(* Logix 5000 project; controller R400_500_XLS vendor 1 type 14 code 216 rev 31.11; software revision 31.01; part 22 of 32 *)
(* tags used below, declared in another part *)
   Abort1 : DINT;   // Not Used
   Alarm : SINT;   // Wait 3 seconds
   AlarmAcked : BOOL;   // Alarm has been acked
   bAlrm : BOOL[64];
   CycExcBuffer : UDT_CYCLE;
   CycleSequence : UDT_CYCLE_SEQUENCE;
   DrnSmp : DINT;
   DRYING : DINT;   // Drying id number
   F1rinse : DINT;   // Not Used
   F2rinse : DINT;   // Not Used
   F3rinse : DINT;   // Not Used
   F4rinse : INT;   // Transition for the conductivity based evalutaion
   F4rinse_Tran : INT;   // Transitions for the conductivity based evaluation
   FINAL_RINSE_MAX_NBR : INT;   // Maximum nimber of final rinse
   M : DINT[5];   // Memory Bits
   NbFinalRinseDone : DINT;
   ONS_FC08 : DINT;
   Run : DINT;
   SumpWaterVolume : DINT;   // Sump Water Volume 0 =Low 1= High
   Tmr : TIMER[107];
   WaterSaved : BOOL;   // Water Saved In Sump (Last Final Rinse Water)
   ENABLE : BOOL;   // Enable bit
   FinalRinseCond : REAL;
   I_Pw_Tnk_Lvl_Sw : BOOL;   // Pure water tank level switch
   TreatmentPtr : DINT;
   Unit : Hrdwre;   // Unit Configuration
(* MainProgram, continued *)

ROUTINE WSH_16_TRT_FRINSE   (* ladder *)
// This routine performs the Final Rinse treatments
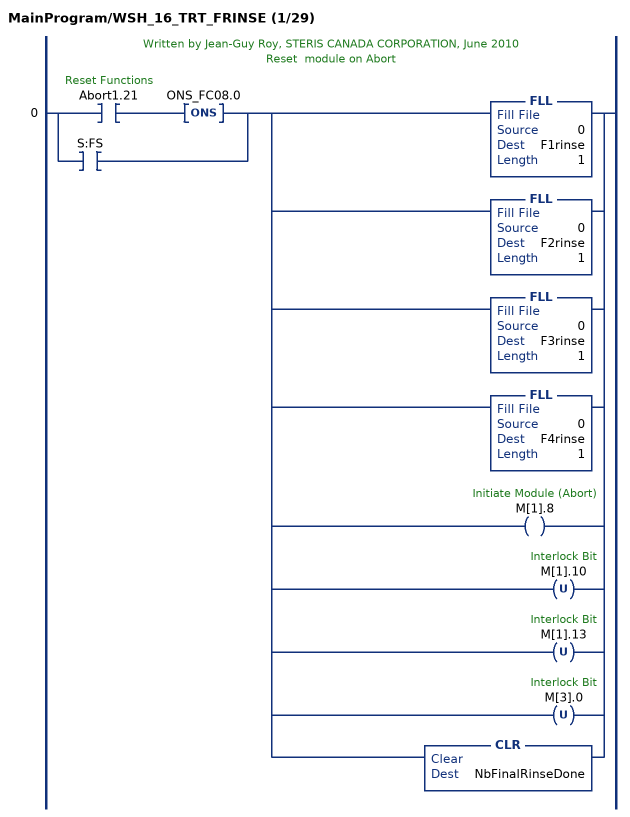
   // Written by Jean-Guy Roy, STERIS CANADA CORPORATION, June 2010
   // Reset  module on Abort
   0: [XIC(Abort1.21) ONS(ONS_FC08.0) ,XIC(S:FS) ][FLL(0,F1rinse,1) ,FLL(0,F2rinse,1) ,FLL(0,F3rinse,1) ,FLL(0,F4rinse,1) ,OTE(M[1].8) ,OTU(M[1].10) ,OTU(M[1].13) ,OTU(M[3].0) ,CLR(NbFinalRinseDone) ];
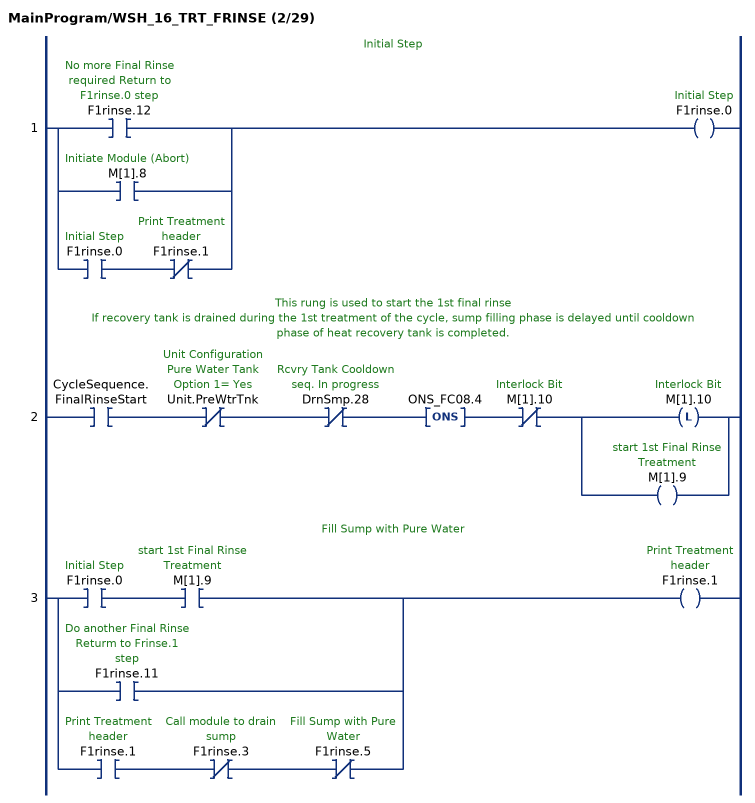
   // Initial Step
   1: [XIC(F1rinse.12) ,XIC(M[1].8) ,XIC(F1rinse.0) XIO(F1rinse.1) ]OTE(F1rinse.0);
   // This rung is used to start the 1st final rinse
   // If recovery tank is drained during the 1st treatment of the cycle, sump filling phase is delayed until cooldown phase of heat recovery tank is completed.
   2: XIC(CycleSequence.FinalRinseStart)XIO(Unit.PreWtrTnk)XIO(DrnSmp.28)ONS(ONS_FC08.4)XIO(M[1].10)[OTL(M[1].10) ,OTE(M[1].9) ];
   // Fill Sump with Pure Water
   3: [XIC(F1rinse.0) XIC(M[1].9) ,XIC(F1rinse.11) ,XIC(F1rinse.1) XIO(F1rinse.3) XIO(F1rinse.5) ]OTE(F1rinse.1);
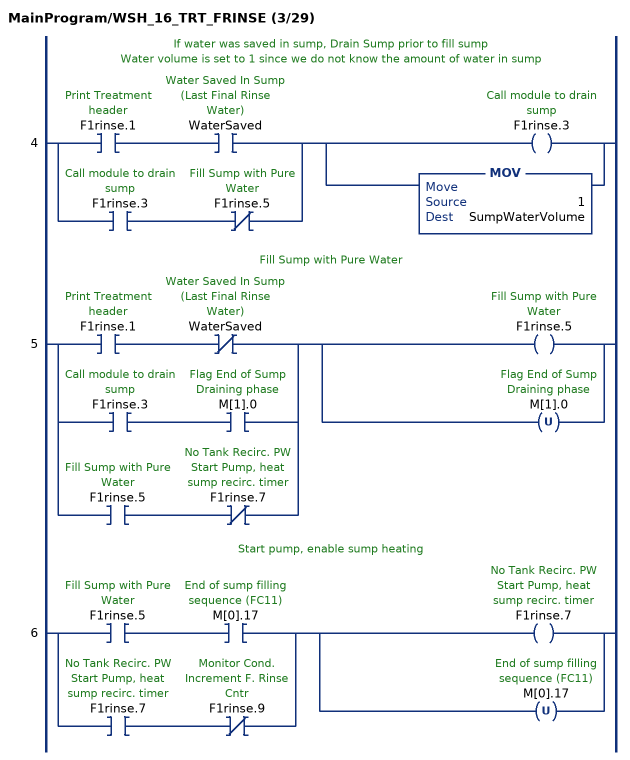
   // If water was saved in sump, Drain Sump prior to fill sump
   // Water volume is set to 1 since we do not know the amount of water in sump
   4: [XIC(F1rinse.1) XIC(WaterSaved) ,XIC(F1rinse.3) XIO(F1rinse.5) ][OTE(F1rinse.3) ,MOV(1,SumpWaterVolume) ];
   // Fill Sump with Pure Water
   5: [[XIC(F1rinse.1) XIO(WaterSaved) ,XIC(F1rinse.3) XIC(M[1].0) ] ,XIC(F1rinse.5) XIO(F1rinse.7) ][OTE(F1rinse.5) ,OTU(M[1].0) ];
   // Start pump, enable sump heating
   6: [XIC(F1rinse.5) XIC(M[0].17) ,XIC(F1rinse.7) XIO(F1rinse.9) ][OTE(F1rinse.7) ,OTU(M[0].17) ];
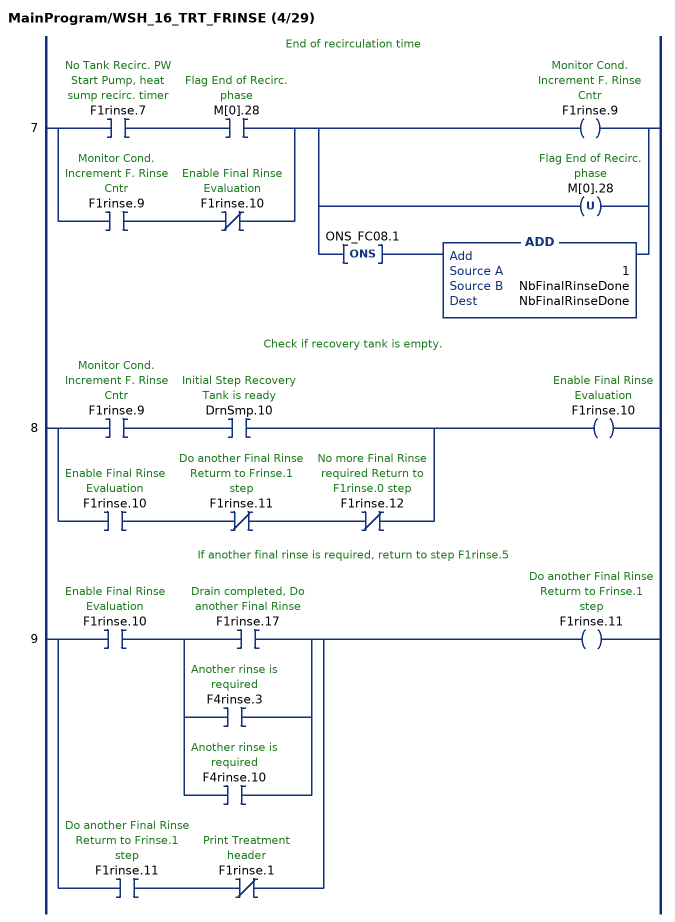
   // End of recirculation time
   7: [XIC(F1rinse.7) XIC(M[0].28) ,XIC(F1rinse.9) XIO(F1rinse.10) ][[OTE(F1rinse.9) ,OTU(M[0].28) ] ,ONS(ONS_FC08.1) ADD(1,NbFinalRinseDone,NbFinalRinseDone) ];
   // Check if recovery tank is empty.
   8: [XIC(F1rinse.9) XIC(DrnSmp.10) ,XIC(F1rinse.10) XIO(F1rinse.11) XIO(F1rinse.12) ]OTE(F1rinse.10);
   // If another final rinse is required, return to step F1rinse.5
   9: [XIC(F1rinse.10) [XIC(F1rinse.17) ,XIC(F4rinse.3) ,XIC(F4rinse.10) ] ,XIC(F1rinse.11) XIO(F1rinse.1) ]OTE(F1rinse.11);
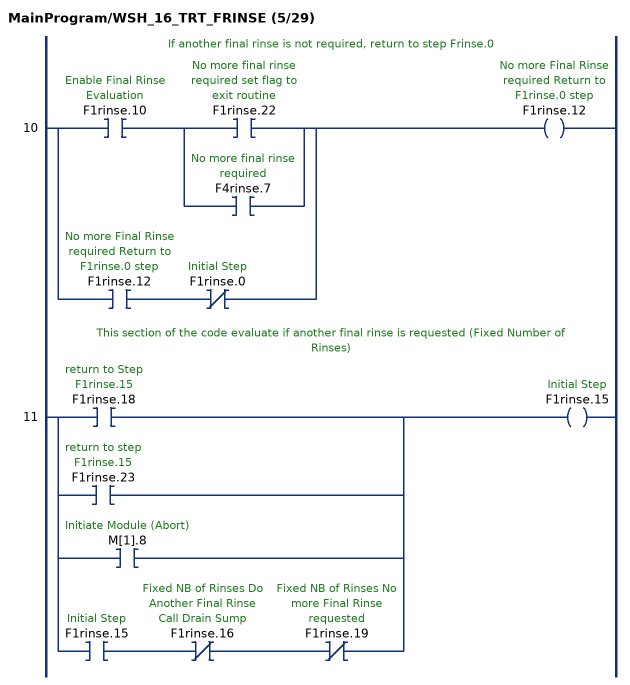
   // If another final rinse is not required, return to step Frinse.0
   10: [XIC(F1rinse.10) [XIC(F1rinse.22) ,XIC(F4rinse.7) ] ,XIC(F1rinse.12) XIO(F1rinse.0) ]OTE(F1rinse.12);
   // This section of the code evaluate if another final rinse is requested (Fixed Number of Rinses)
   11: [XIC(F1rinse.18) ,XIC(F1rinse.23) ,XIC(M[1].8) ,XIC(F1rinse.15) XIO(F1rinse.16) XIO(F1rinse.19) ]OTE(F1rinse.15);
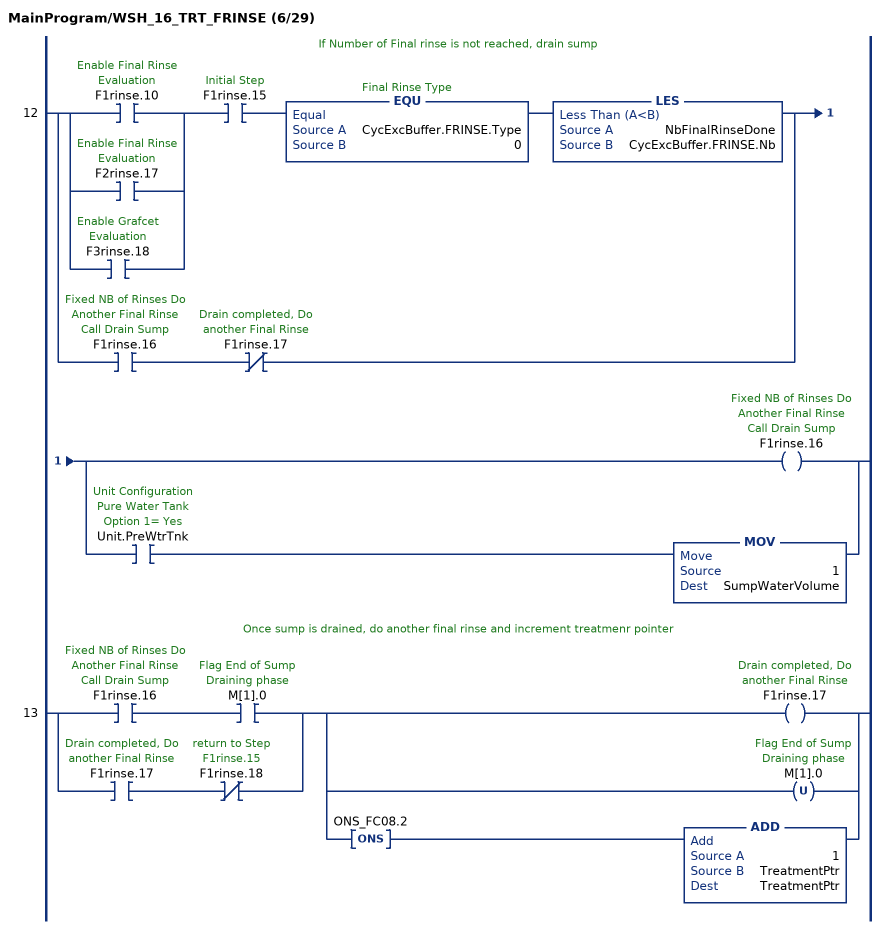
   // If Number of Final rinse is not reached, drain sump
   12: [[XIC(F1rinse.10) ,XIC(F2rinse.17) ,XIC(F3rinse.18) ] XIC(F1rinse.15) EQU(CycExcBuffer.FRINSE.Type,0) LES(NbFinalRinseDone,CycExcBuffer.FRINSE.Nb) ,XIC(F1rinse.16) XIO(F1rinse.17) ][OTE(F1rinse.16) ,XIC(Unit.PreWtrTnk) MOV(1,SumpWaterVolume) ];
   // Once sump is drained, do another final rinse and increment treatmenr pointer
   13: [XIC(F1rinse.16) XIC(M[1].0) ,XIC(F1rinse.17) XIO(F1rinse.18) ][OTE(F1rinse.17) ,OTU(M[1].0) ,ONS(ONS_FC08.2) ADD(1,TreatmentPtr,TreatmentPtr) ];
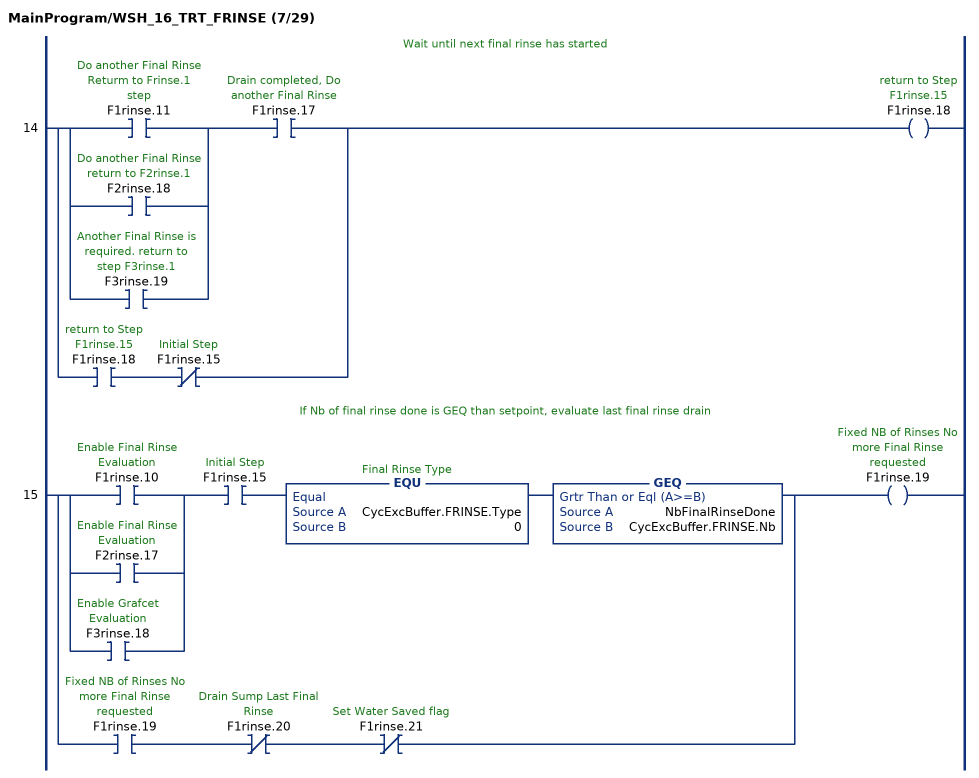
   // Wait until next final rinse has started
   14: [[XIC(F1rinse.11) ,XIC(F2rinse.18) ,XIC(F3rinse.19) ] XIC(F1rinse.17) ,XIC(F1rinse.18) XIO(F1rinse.15) ]OTE(F1rinse.18);
   // If Nb of final rinse done is GEQ than setpoint, evaluate last final rinse drain
   15: [[XIC(F1rinse.10) ,XIC(F2rinse.17) ,XIC(F3rinse.18) ] XIC(F1rinse.15) EQU(CycExcBuffer.FRINSE.Type,0) GEQ(NbFinalRinseDone,CycExcBuffer.FRINSE.Nb) ,XIC(F1rinse.19) XIO(F1rinse.20) XIO(F1rinse.21) ]OTE(F1rinse.19);
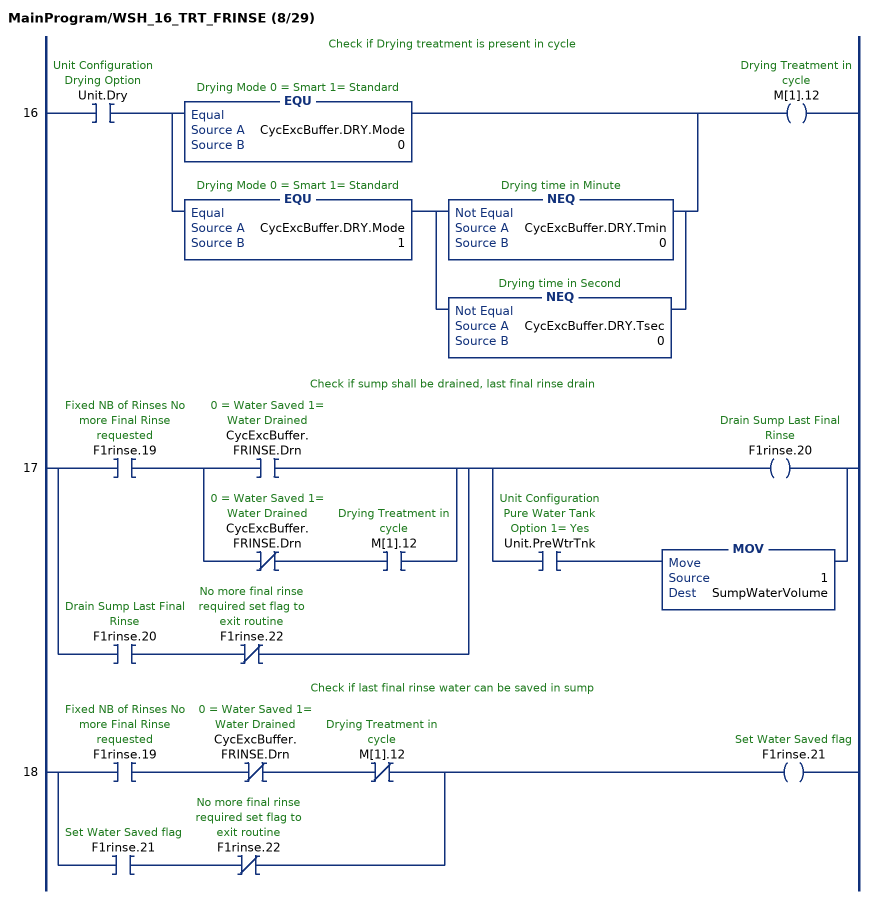
   // Check if Drying treatment is present in cycle
   16: XIC(Unit.Dry)[EQU(CycExcBuffer.DRY.Mode,0) ,EQU(CycExcBuffer.DRY.Mode,1) [NEQ(CycExcBuffer.DRY.Tmin,0) ,NEQ(CycExcBuffer.DRY.Tsec,0) ] ]OTE(M[1].12);
   // Check if sump shall be drained, last final rinse drain
   17: [XIC(F1rinse.19) [XIC(CycExcBuffer.FRINSE.Drn) ,XIO(CycExcBuffer.FRINSE.Drn) XIC(M[1].12) ] ,XIC(F1rinse.20) XIO(F1rinse.22) ][OTE(F1rinse.20) ,XIC(Unit.PreWtrTnk) MOV(1,SumpWaterVolume) ];
   // Check if last final rinse water can be saved in sump
   18: [XIC(F1rinse.19) XIO(CycExcBuffer.FRINSE.Drn) XIO(M[1].12) ,XIC(F1rinse.21) XIO(F1rinse.22) ]OTE(F1rinse.21);
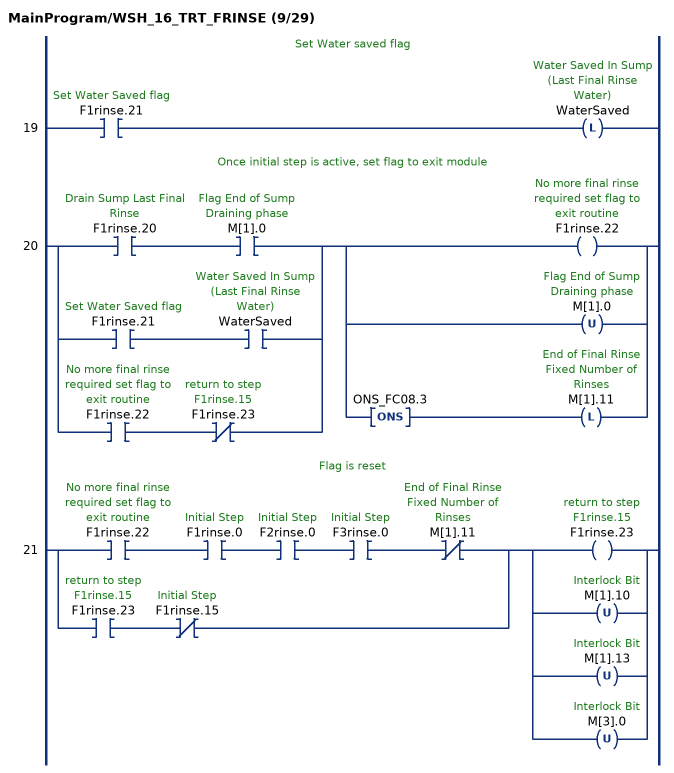
   // Set Water saved flag
   19: XIC(F1rinse.21)OTL(WaterSaved);
   // Once initial step is active, set flag to exit module
   20: [XIC(F1rinse.20) XIC(M[1].0) ,XIC(F1rinse.21) XIC(WaterSaved) ,XIC(F1rinse.22) XIO(F1rinse.23) ][OTE(F1rinse.22) ,OTU(M[1].0) ,ONS(ONS_FC08.3) OTL(M[1].11) ];
   // Flag is reset
   21: [XIC(F1rinse.22) XIC(F1rinse.0) XIC(F2rinse.0) XIC(F3rinse.0) XIO(M[1].11) ,XIC(F1rinse.23) XIO(F1rinse.15) ][OTE(F1rinse.23) ,OTU(M[1].10) ,OTU(M[1].13) ,OTU(M[3].0) ];
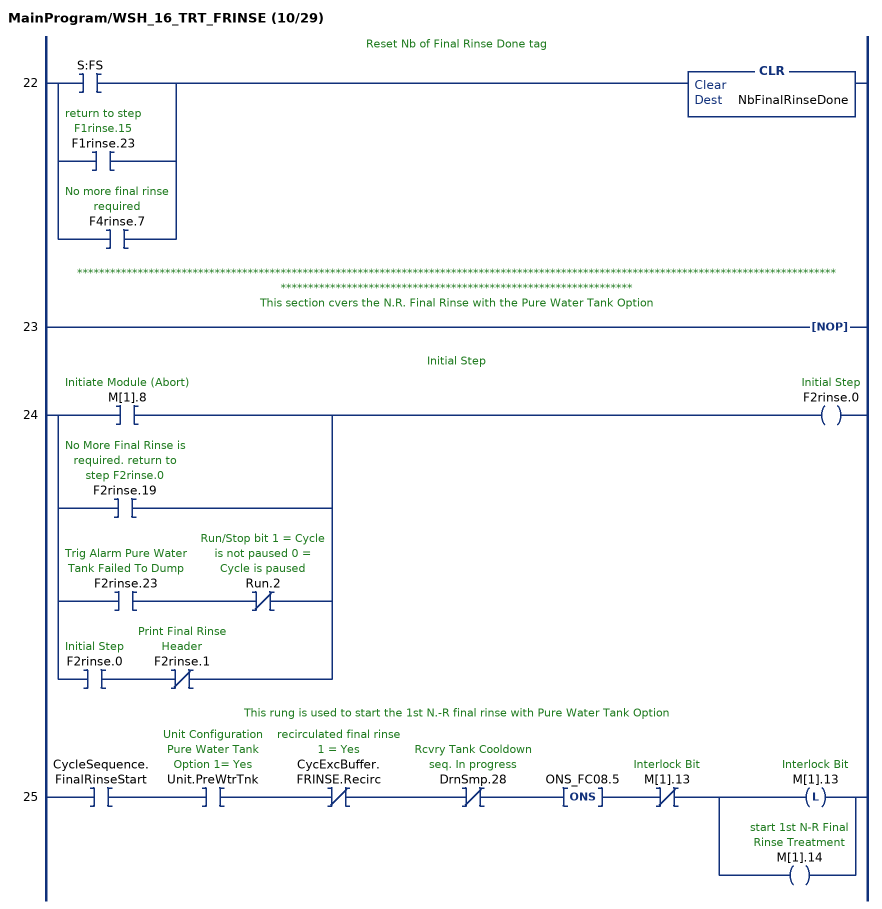
   // Reset Nb of Final Rinse Done tag
   22: [XIC(S:FS) ,XIC(F1rinse.23) ,XIC(F4rinse.7) ]CLR(NbFinalRinseDone);
   // **********************************************************************************************************************************************************************************************************
   // This section cvers the N.R. Final Rinse with the Pure Water Tank Option
   23: NOP();
   // Initial Step
   24: [XIC(M[1].8) ,XIC(F2rinse.19) ,XIC(F2rinse.23) XIO(Run.2) ,XIC(F2rinse.0) XIO(F2rinse.1) ]OTE(F2rinse.0);
   // This rung is used to start the 1st N.-R final rinse with Pure Water Tank Option
   25: XIC(CycleSequence.FinalRinseStart)XIC(Unit.PreWtrTnk)XIO(CycExcBuffer.FRINSE.Recirc)XIO(DrnSmp.28)ONS(ONS_FC08.5)XIO(M[1].13)[OTL(M[1].13) ,OTE(M[1].14) ];
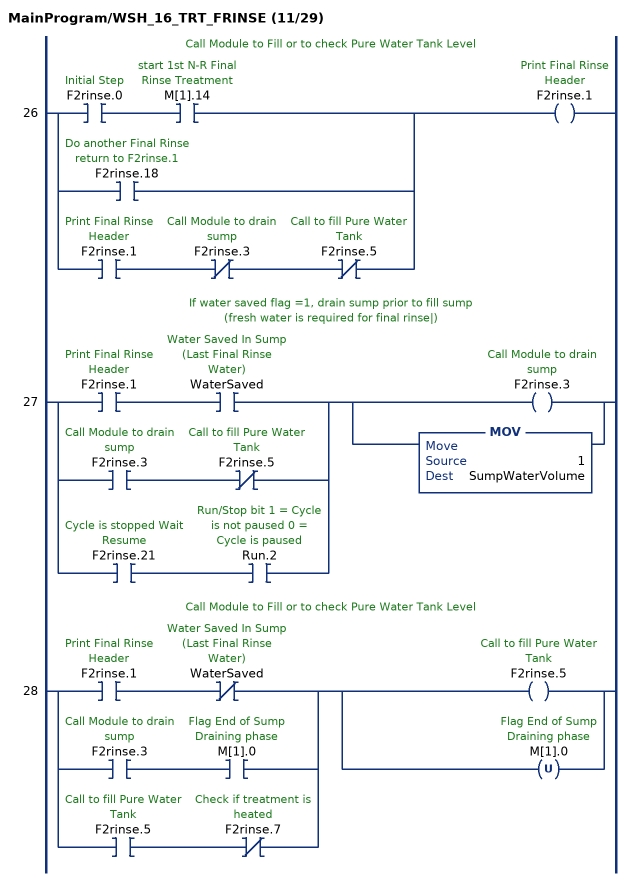
   // Call Module to Fill or to check Pure Water Tank Level
   26: [XIC(F2rinse.0) XIC(M[1].14) ,XIC(F2rinse.18) ,XIC(F2rinse.1) XIO(F2rinse.3) XIO(F2rinse.5) ]OTE(F2rinse.1);
   // If water saved flag =1, drain sump prior to fill sump
   // (fresh water is required for final rinse|)
   27: [XIC(F2rinse.1) XIC(WaterSaved) ,XIC(F2rinse.3) XIO(F2rinse.5) ,XIC(F2rinse.21) XIC(Run.2) ][OTE(F2rinse.3) ,MOV(1,SumpWaterVolume) ];
   // Call Module to Fill or to check Pure Water Tank Level
   28: [XIC(F2rinse.1) XIO(WaterSaved) ,XIC(F2rinse.3) XIC(M[1].0) ,XIC(F2rinse.5) XIO(F2rinse.7) ][OTE(F2rinse.5) ,OTU(M[1].0) ];
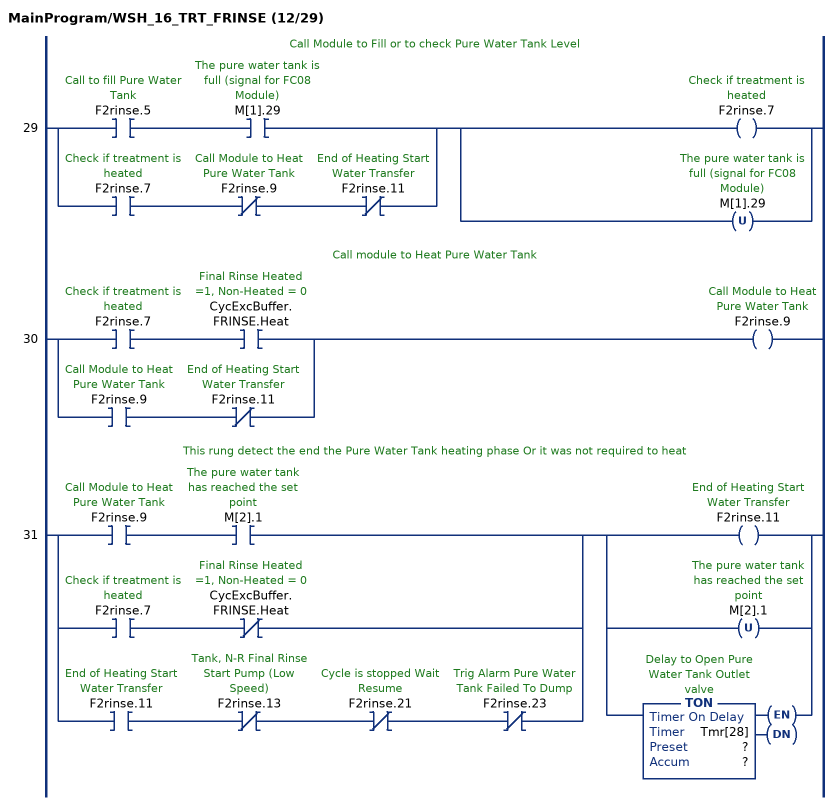
   // Call Module to Fill or to check Pure Water Tank Level
   29: [XIC(F2rinse.5) XIC(M[1].29) ,XIC(F2rinse.7) XIO(F2rinse.9) XIO(F2rinse.11) ][OTE(F2rinse.7) ,OTU(M[1].29) ];
   // Call module to Heat Pure Water Tank
   30: [XIC(F2rinse.7) XIC(CycExcBuffer.FRINSE.Heat) ,XIC(F2rinse.9) XIO(F2rinse.11) ]OTE(F2rinse.9);
   // This rung detect the end the Pure Water Tank heating phase Or it was not required to heat
   31: [XIC(F2rinse.9) XIC(M[2].1) ,XIC(F2rinse.7) XIO(CycExcBuffer.FRINSE.Heat) ,XIC(F2rinse.11) XIO(F2rinse.13) XIO(F2rinse.21) XIO(F2rinse.23) ][OTE(F2rinse.11) ,OTU(M[2].1) ,TON(Tmr[28],?,?) ];
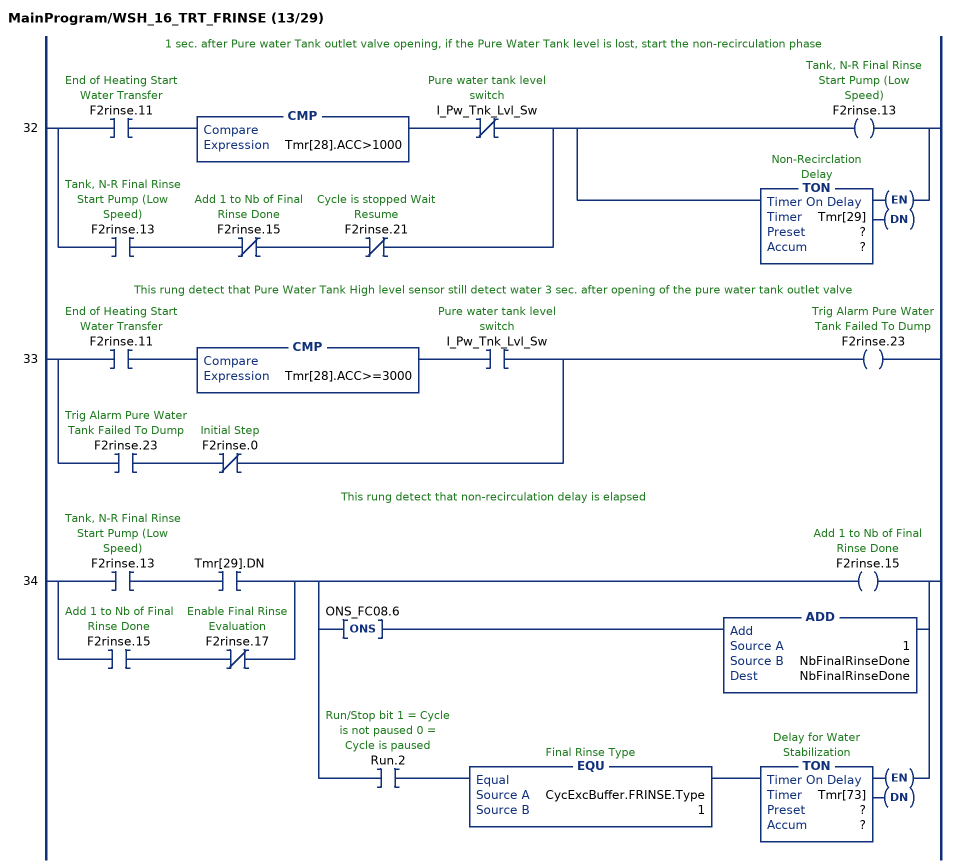
   // 1 sec. after Pure water Tank outlet valve opening, if the Pure Water Tank level is lost, start the non-recirculation phase
   32: [XIC(F2rinse.11) CMP(Tmr[28].ACC>1000) XIO(I_Pw_Tnk_Lvl_Sw) ,XIC(F2rinse.13) XIO(F2rinse.15) XIO(F2rinse.21) ][OTE(F2rinse.13) ,TON(Tmr[29],?,?) ];
   // This rung detect that Pure Water Tank High level sensor still detect water 3 sec. after opening of the pure water tank outlet valve
   33: [XIC(F2rinse.11) CMP(Tmr[28].ACC>=3000) XIC(I_Pw_Tnk_Lvl_Sw) ,XIC(F2rinse.23) XIO(F2rinse.0) ]OTE(F2rinse.23);
   // This rung detect that non-recirculation delay is elapsed
   34: [XIC(F2rinse.13) XIC(Tmr[29].DN) ,XIC(F2rinse.15) XIO(F2rinse.17) ][OTE(F2rinse.15) ,ONS(ONS_FC08.6) ADD(1,NbFinalRinseDone,NbFinalRinseDone) ,XIC(Run.2) EQU(CycExcBuffer.FRINSE.Type,1) TON(Tmr[73],?,?) ];
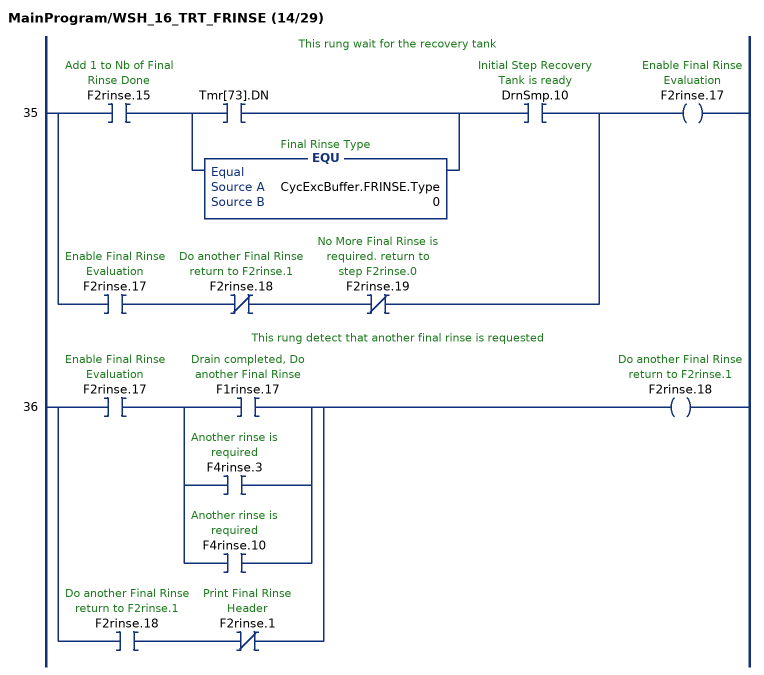
   // This rung wait for the recovery tank
   35: [XIC(F2rinse.15) [XIC(Tmr[73].DN) ,EQU(CycExcBuffer.FRINSE.Type,0) ] XIC(DrnSmp.10) ,XIC(F2rinse.17) XIO(F2rinse.18) XIO(F2rinse.19) ]OTE(F2rinse.17);
   // This rung detect that another final rinse is requested
   36: [XIC(F2rinse.17) [XIC(F1rinse.17) ,XIC(F4rinse.3) ,XIC(F4rinse.10) ] ,XIC(F2rinse.18) XIO(F2rinse.1) ]OTE(F2rinse.18);
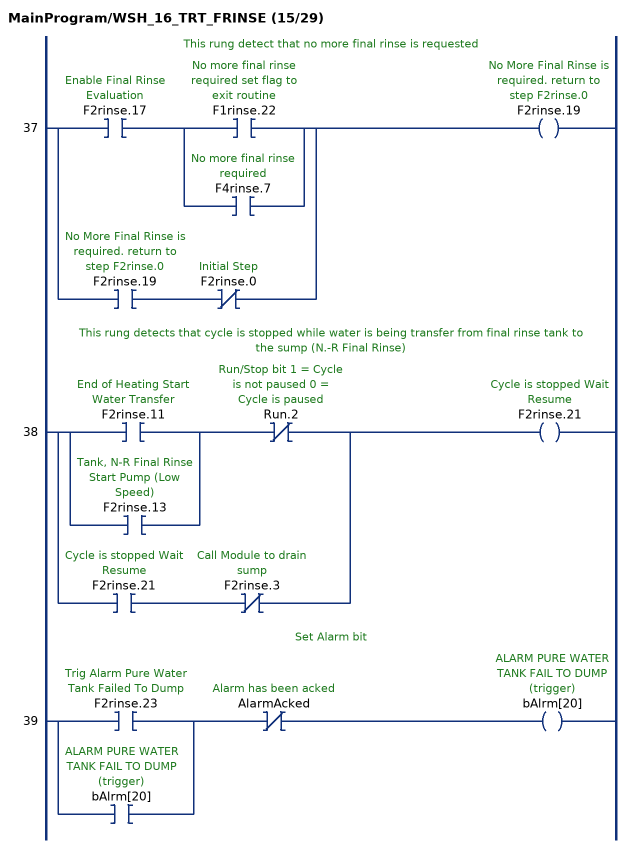
   // This rung detect that no more final rinse is requested
   37: [XIC(F2rinse.17) [XIC(F1rinse.22) ,XIC(F4rinse.7) ] ,XIC(F2rinse.19) XIO(F2rinse.0) ]OTE(F2rinse.19);
   // This rung detects that cycle is stopped while water is being transfer from final rinse tank to the sump (N.-R Final Rinse)
   38: [[XIC(F2rinse.11) ,XIC(F2rinse.13) ] XIO(Run.2) ,XIC(F2rinse.21) XIO(F2rinse.3) ]OTE(F2rinse.21);
   // Set Alarm bit
   39: [XIC(F2rinse.23) ,XIC(bAlrm[20]) ]XIO(AlarmAcked)OTE(bAlrm[20]);
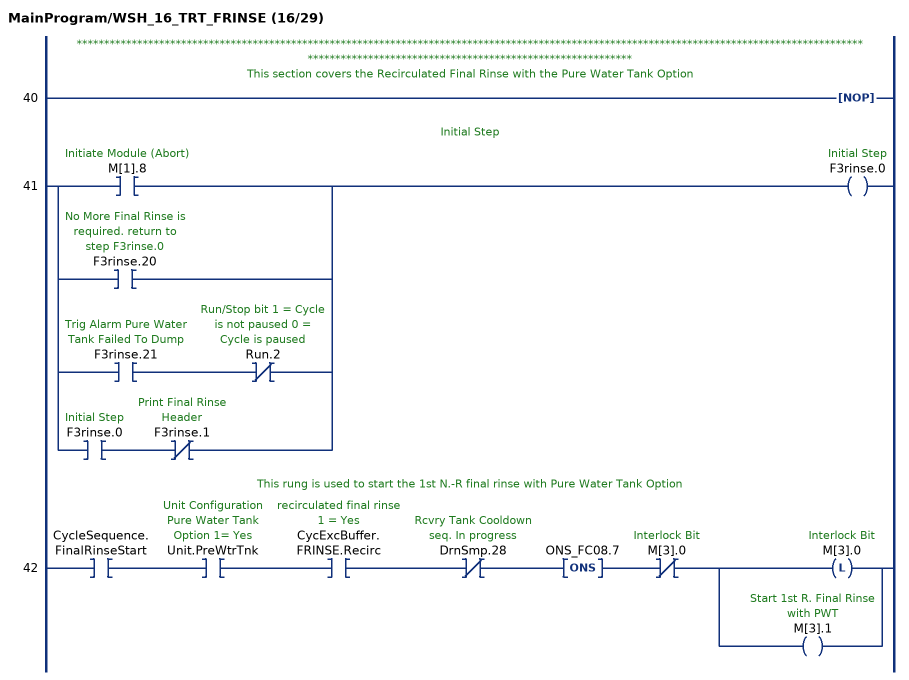
   // **********************************************************************************************************************************************************************************************************
   // This section covers the Recirculated Final Rinse with the Pure Water Tank Option
   40: NOP();
   // Initial Step
   41: [XIC(M[1].8) ,XIC(F3rinse.20) ,XIC(F3rinse.21) XIO(Run.2) ,XIC(F3rinse.0) XIO(F3rinse.1) ]OTE(F3rinse.0);
   // This rung is used to start the 1st N.-R final rinse with Pure Water Tank Option
   42: XIC(CycleSequence.FinalRinseStart)XIC(Unit.PreWtrTnk)XIC(CycExcBuffer.FRINSE.Recirc)XIO(DrnSmp.28)ONS(ONS_FC08.7)XIO(M[3].0)[OTL(M[3].0) ,OTE(M[3].1) ];
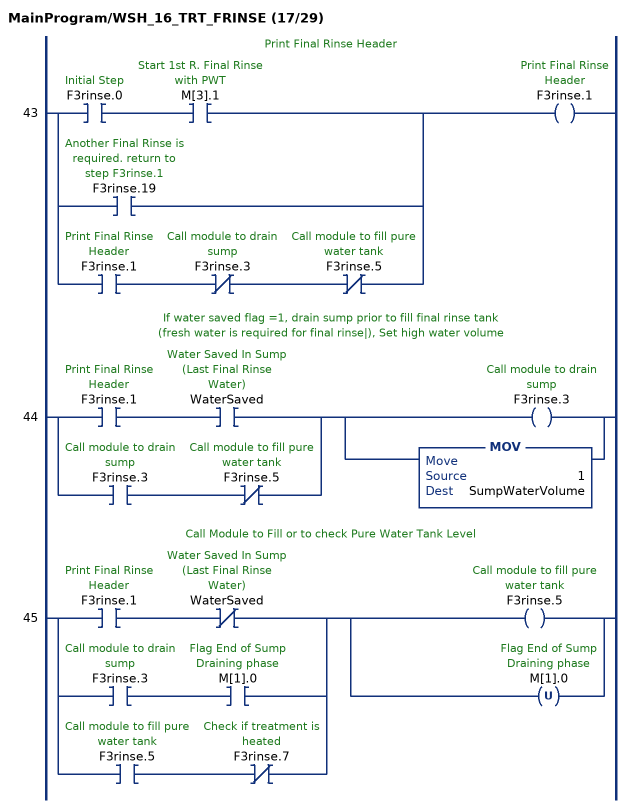
   // Print Final Rinse Header
   43: [XIC(F3rinse.0) XIC(M[3].1) ,XIC(F3rinse.19) ,XIC(F3rinse.1) XIO(F3rinse.3) XIO(F3rinse.5) ]OTE(F3rinse.1);
   // If water saved flag =1, drain sump prior to fill final rinse tank
   // (fresh water is required for final rinse|), Set high water volume
   44: [XIC(F3rinse.1) XIC(WaterSaved) ,XIC(F3rinse.3) XIO(F3rinse.5) ][OTE(F3rinse.3) ,MOV(1,SumpWaterVolume) ];
   // Call Module to Fill or to check Pure Water Tank Level
   45: [XIC(F3rinse.1) XIO(WaterSaved) ,XIC(F3rinse.3) XIC(M[1].0) ,XIC(F3rinse.5) XIO(F3rinse.7) ][OTE(F3rinse.5) ,OTU(M[1].0) ];
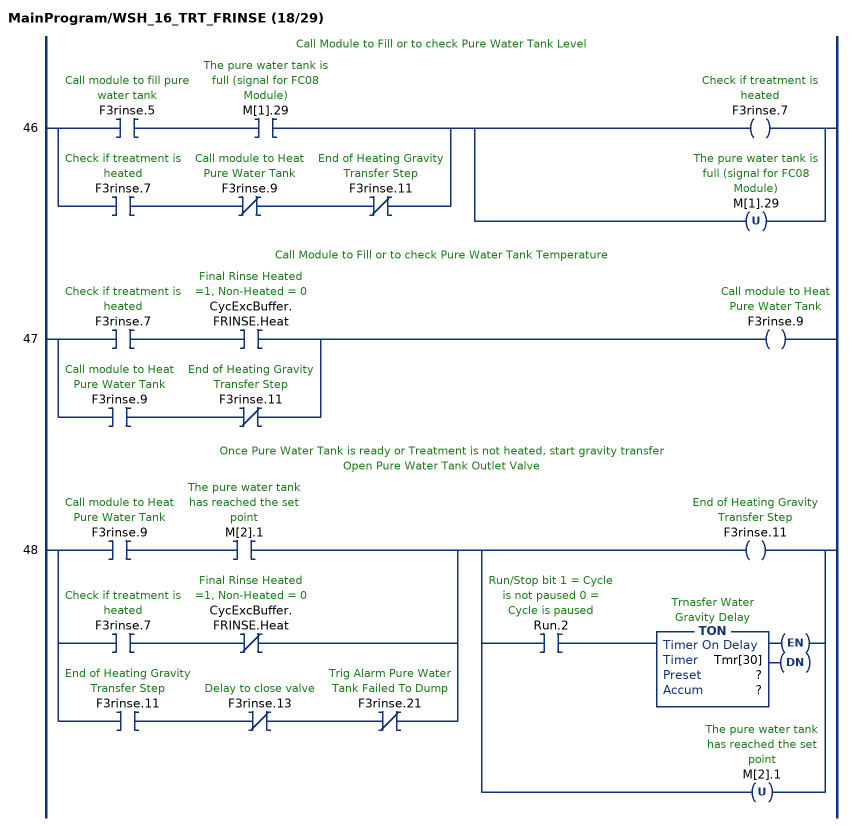
   // Call Module to Fill or to check Pure Water Tank Level
   46: [XIC(F3rinse.5) XIC(M[1].29) ,XIC(F3rinse.7) XIO(F3rinse.9) XIO(F3rinse.11) ][OTE(F3rinse.7) ,OTU(M[1].29) ];
   // Call Module to Fill or to check Pure Water Tank Temperature
   47: [XIC(F3rinse.7) XIC(CycExcBuffer.FRINSE.Heat) ,XIC(F3rinse.9) XIO(F3rinse.11) ]OTE(F3rinse.9);
   // Once Pure Water Tank is ready or Treatment is not heated, start gravity transfer
   // Open Pure Water Tank Outlet Valve
   48: [XIC(F3rinse.9) XIC(M[2].1) ,XIC(F3rinse.7) XIO(CycExcBuffer.FRINSE.Heat) ,XIC(F3rinse.11) XIO(F3rinse.13) XIO(F3rinse.21) ][OTE(F3rinse.11) ,XIC(Run.2) TON(Tmr[30],?,?) ,OTU(M[2].1) ];
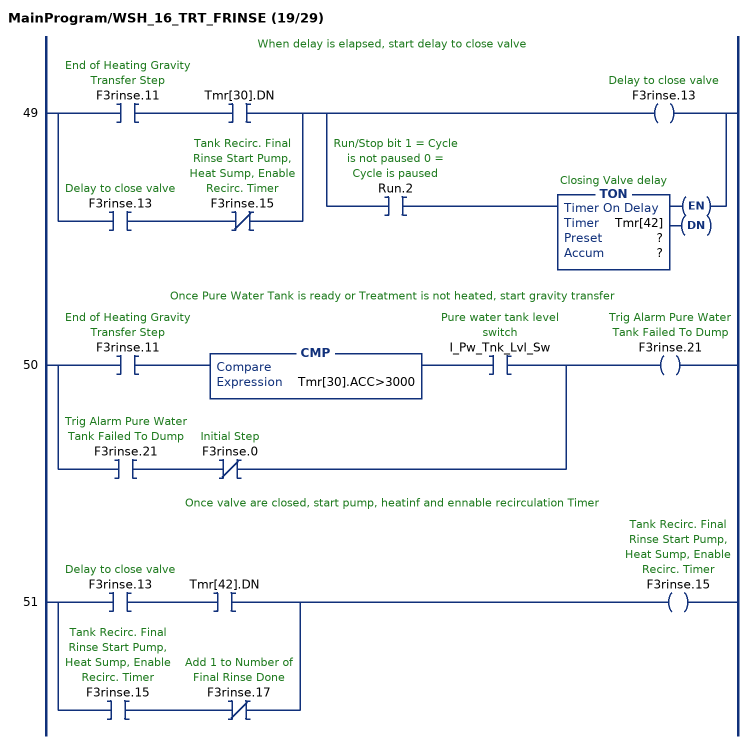
   // When delay is elapsed, start delay to close valve
   49: [XIC(F3rinse.11) XIC(Tmr[30].DN) ,XIC(F3rinse.13) XIO(F3rinse.15) ][OTE(F3rinse.13) ,XIC(Run.2) TON(Tmr[42],?,?) ];
   // Once Pure Water Tank is ready or Treatment is not heated, start gravity transfer
   50: [XIC(F3rinse.11) CMP(Tmr[30].ACC>3000) XIC(I_Pw_Tnk_Lvl_Sw) ,XIC(F3rinse.21) XIO(F3rinse.0) ]OTE(F3rinse.21);
   // Once valve are closed, start pump, heatinf and ennable recirculation Timer
   51: [XIC(F3rinse.13) XIC(Tmr[42].DN) ,XIC(F3rinse.15) XIO(F3rinse.17) ]OTE(F3rinse.15);
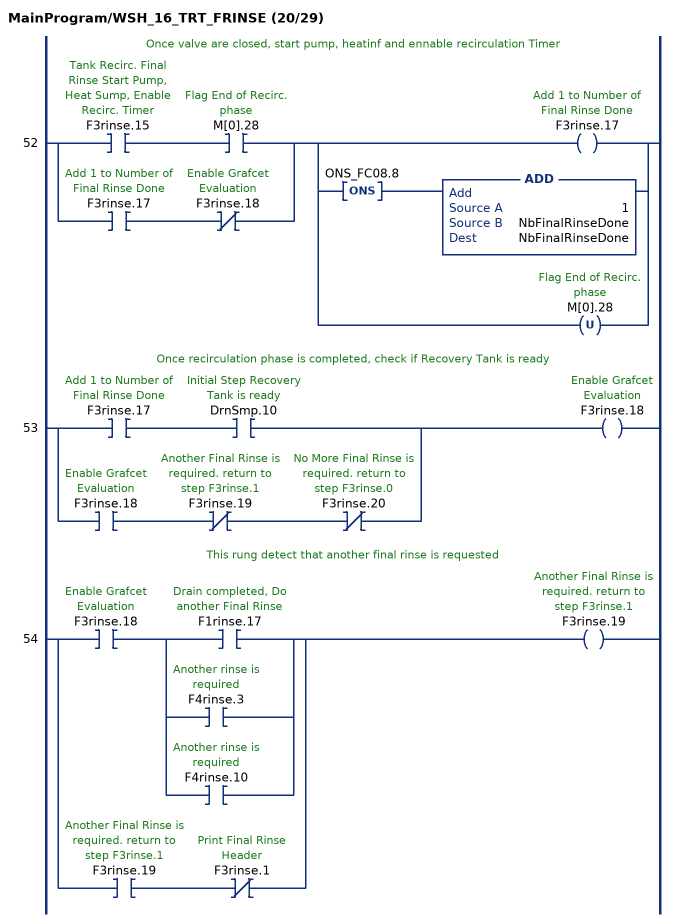
   // Once valve are closed, start pump, heatinf and ennable recirculation Timer
   52: [XIC(F3rinse.15) XIC(M[0].28) ,XIC(F3rinse.17) XIO(F3rinse.18) ][OTE(F3rinse.17) ,ONS(ONS_FC08.8) ADD(1,NbFinalRinseDone,NbFinalRinseDone) ,OTU(M[0].28) ];
   // Once recirculation phase is completed, check if Recovery Tank is ready
   53: [XIC(F3rinse.17) XIC(DrnSmp.10) ,XIC(F3rinse.18) XIO(F3rinse.19) XIO(F3rinse.20) ]OTE(F3rinse.18);
   // This rung detect that another final rinse is requested
   54: [XIC(F3rinse.18) [XIC(F1rinse.17) ,XIC(F4rinse.3) ,XIC(F4rinse.10) ] ,XIC(F3rinse.19) XIO(F3rinse.1) ]OTE(F3rinse.19);
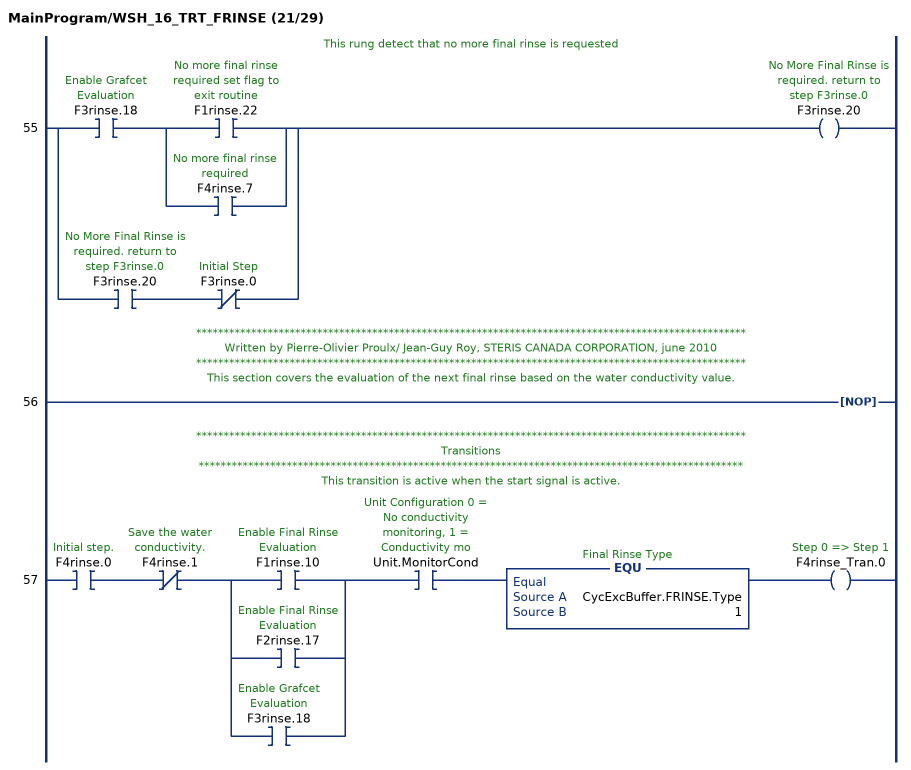
   // This rung detect that no more final rinse is requested
   55: [XIC(F3rinse.18) [XIC(F1rinse.22) ,XIC(F4rinse.7) ] ,XIC(F3rinse.20) XIO(F3rinse.0) ]OTE(F3rinse.20);
   // ****************************************************************************************************
   // Written by Pierre-Olivier Proulx/ Jean-Guy Roy, STERIS CANADA CORPORATION, june 2010
   // ****************************************************************************************************
   // This section covers the evaluation of the next final rinse based on the water conductivity value.
   56: NOP();
   // ****************************************************************************************************
   // Transitions
   // ***************************************************************************************************
   // This transition is active when the start signal is active.
   57: XIC(F4rinse.0)XIO(F4rinse.1)[XIC(F1rinse.10) ,XIC(F2rinse.17) ,XIC(F3rinse.18) ]XIC(Unit.MonitorCond)EQU(CycExcBuffer.FRINSE.Type,1)OTE(F4rinse_Tran.0);
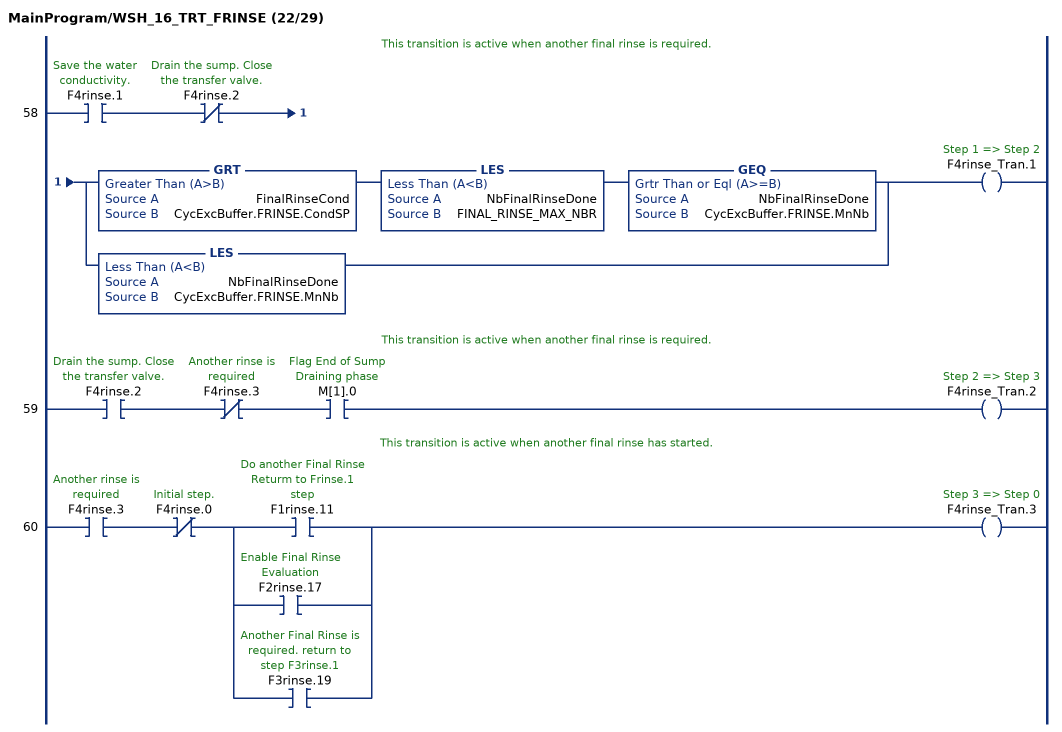
   // This transition is active when another final rinse is required.
   58: XIC(F4rinse.1)XIO(F4rinse.2)[GRT(FinalRinseCond,CycExcBuffer.FRINSE.CondSP) LES(NbFinalRinseDone,FINAL_RINSE_MAX_NBR) GEQ(NbFinalRinseDone,CycExcBuffer.FRINSE.MnNb) ,LES(NbFinalRinseDone,CycExcBuffer.FRINSE.MnNb) ]OTE(F4rinse_Tran.1);
   // This transition is active when another final rinse is required.
   59: XIC(F4rinse.2)XIO(F4rinse.3)XIC(M[1].0)OTE(F4rinse_Tran.2);
   // This transition is active when another final rinse has started.
   60: XIC(F4rinse.3)XIO(F4rinse.0)[XIC(F1rinse.11) ,XIC(F2rinse.17) ,XIC(F3rinse.19) ]OTE(F4rinse_Tran.3);
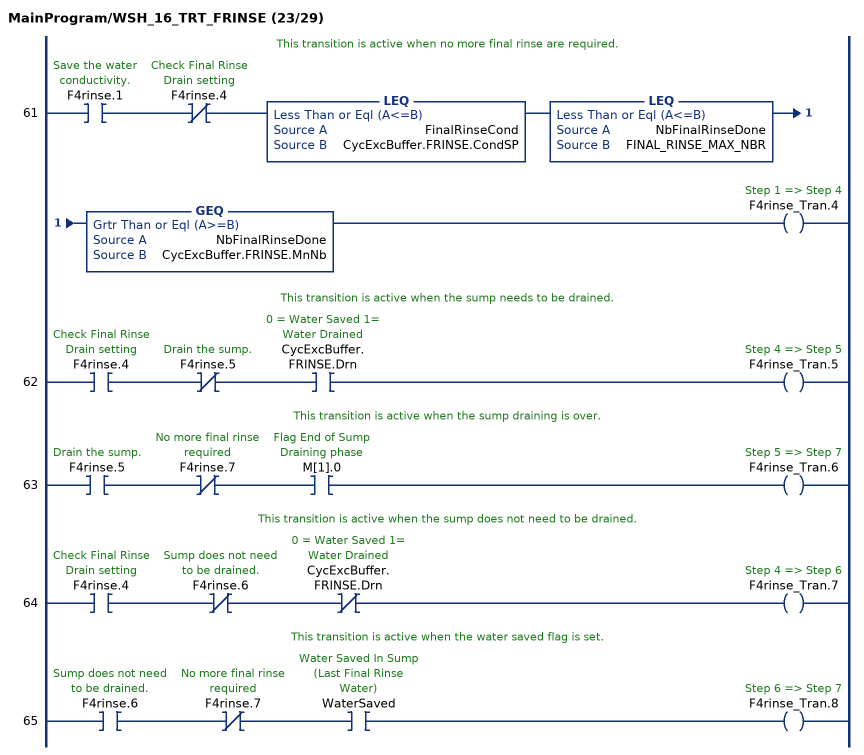
   // This transition is active when no more final rinse are required.
   61: XIC(F4rinse.1)XIO(F4rinse.4)LEQ(FinalRinseCond,CycExcBuffer.FRINSE.CondSP)LEQ(NbFinalRinseDone,FINAL_RINSE_MAX_NBR)GEQ(NbFinalRinseDone,CycExcBuffer.FRINSE.MnNb)OTE(F4rinse_Tran.4);
   // This transition is active when the sump needs to be drained.
   62: XIC(F4rinse.4)XIO(F4rinse.5)XIC(CycExcBuffer.FRINSE.Drn)OTE(F4rinse_Tran.5);
   // This transition is active when the sump draining is over.
   63: XIC(F4rinse.5)XIO(F4rinse.7)XIC(M[1].0)OTE(F4rinse_Tran.6);
   // This transition is active when the sump does not need to be drained.
   64: XIC(F4rinse.4)XIO(F4rinse.6)XIO(CycExcBuffer.FRINSE.Drn)OTE(F4rinse_Tran.7);
   // This transition is active when the water saved flag is set.
   65: XIC(F4rinse.6)XIO(F4rinse.7)XIC(WaterSaved)OTE(F4rinse_Tran.8);
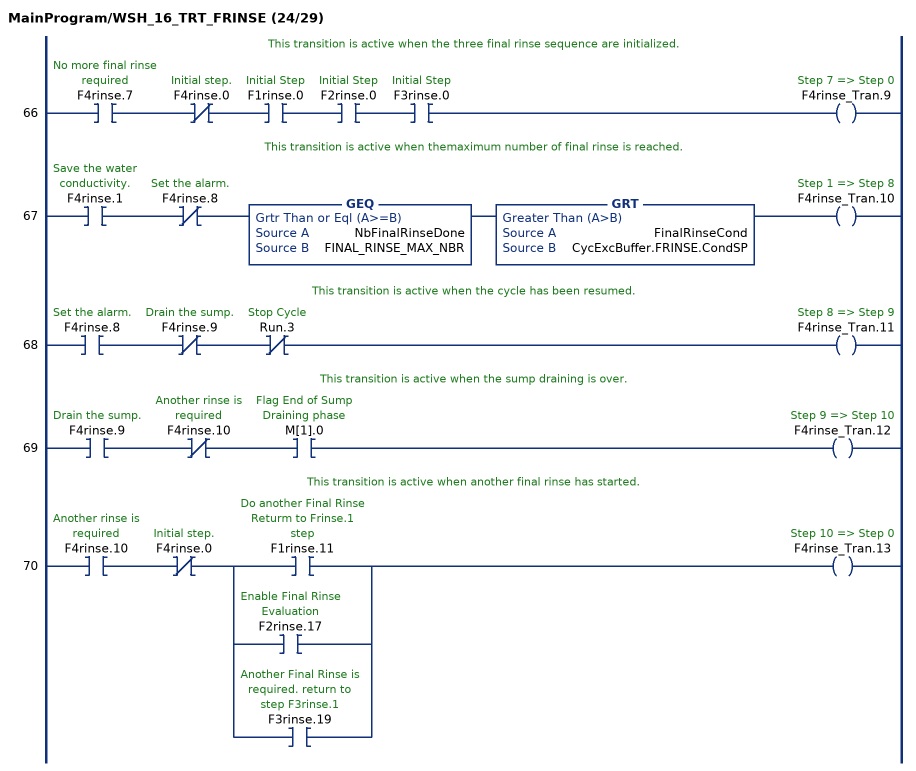
   // This transition is active when the three final rinse sequence are initialized.
   66: XIC(F4rinse.7)XIO(F4rinse.0)XIC(F1rinse.0)XIC(F2rinse.0)XIC(F3rinse.0)OTE(F4rinse_Tran.9);
   // This transition is active when themaximum number of final rinse is reached.
   67: XIC(F4rinse.1)XIO(F4rinse.8)GEQ(NbFinalRinseDone,FINAL_RINSE_MAX_NBR)GRT(FinalRinseCond,CycExcBuffer.FRINSE.CondSP)OTE(F4rinse_Tran.10);
   // This transition is active when the cycle has been resumed.
   68: XIC(F4rinse.8)XIO(F4rinse.9)XIO(Run.3)OTE(F4rinse_Tran.11);
   // This transition is active when the sump draining is over.
   69: XIC(F4rinse.9)XIO(F4rinse.10)XIC(M[1].0)OTE(F4rinse_Tran.12);
   // This transition is active when another final rinse has started.
   70: XIC(F4rinse.10)XIO(F4rinse.0)[XIC(F1rinse.11) ,XIC(F2rinse.17) ,XIC(F3rinse.19) ]OTE(F4rinse_Tran.13);
